SUBAPPLICATION Boot_Melden_OPC (* Station meldet ihren Start an STG1: steigende Flanke von READY ruft die Boot-Methode mit der STG-Nummer auf (ohne VT) *)
  (* Standard: 61499-2; Description: Copyright (c) 2026 Meisterschulen am Ostbahnhof This program and the accompanying materials are made available under the terms of the Eclipse Public License 2.0 which is available at https://www.eclipse.org/legal/epl-2.0/ SPDX-License-Identifier: EPL-2.0 *)
  (* Version 1.1, 2026-10-30, Franz Höpfinger, Meisterschulen am Ostbahnhof, CLIENT_1_0 (Methode) und AX_SUBSCRIBE_1 (READY) je mit Remote_Init_Retry: INITO sofort, nach INITO- (STG1 noch nicht da) neuer Versuch nach 2 s. Vorher hielt die Kette bis 60 s und der Client war danach tot (forte #1092). *)
  (* Version 1.0, 2026-10-29, Franz Höpfinger, Meisterschulen am Ostbahnhof, Neu, Gegenstueck zu Boot_Zaehler_OPC (STG1). AX_SUBSCRIBE_1 startet mit FALSE, daher gibt es nach jedem eigenen Start genau eine steigende Flanke, sobald READY von STG1 ankommt. Reconnect ohne Neustart erzeugt keine Flanke. *)
  PACKAGE MyLib::sys;
  (* Documentation:
  Start an STG1 melden
   Die Station abonniert READY von STG1. Nach dem eigenen Start steht der Wert zunächst auf FALSE; sobald TRUE von STG1 ankommt, ruft die Station einmal die Methode BOOT_MELDUNG mit ihrer Nummer NR auf. STG1 zählt die Starts (Boot_Zaehler_OPC).
  *)
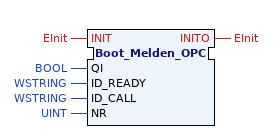
  EVENT_INPUT
    INIT : EInit; (* Initialization Request *)
  END_EVENT
  EVENT_OUTPUT
    INITO : EInit; (* Initialization Confirm *)
  END_EVENT
  VAR_INPUT
    QI : BOOL := TRUE; (* Quality Input - TRUE to enable service *)
    ID_READY : WSTRING; (* Remote-Subscribe READY von STG1 *)
    ID_CALL : WSTRING; (* Remote-Methode BOOT_MELDUNG auf STG1 *)
    NR : UINT; (* Eigene STG-Nummer (2..5) *)
  END_VAR
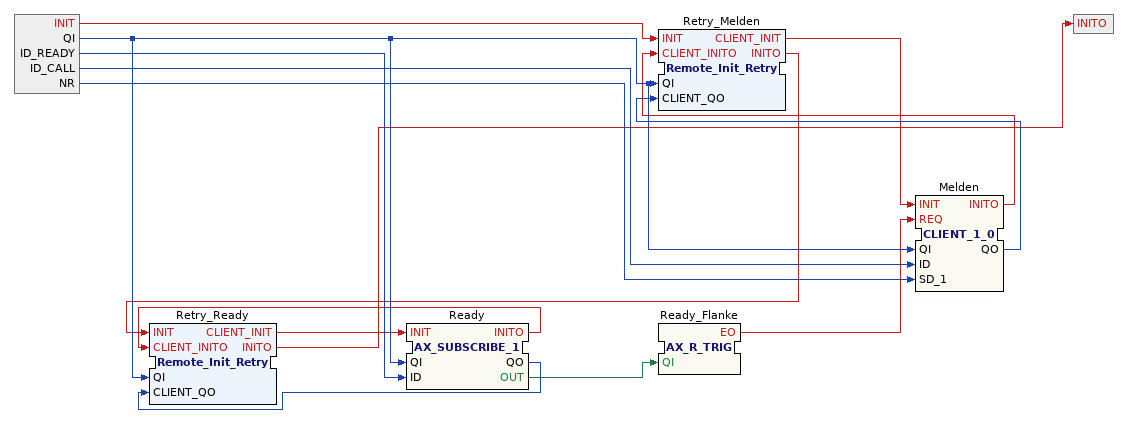
  FBS
    Melden : iec61499::net::CLIENT_1_0;
    Ready : adapter::net::AX_SUBSCRIBE_1;
    Ready_Flanke : adapter::events::unidirectional::AX_R_TRIG;
  END_FBS
  SUBAPPS
    Retry_Melden : MyLib::sys::Remote_Init_Retry;
    Retry_Ready : MyLib::sys::Remote_Init_Retry;
  END_SUBAPPS
  EVENT_CONNECTIONS
    INIT TO Retry_Melden.INIT;
    Retry_Melden.CLIENT_INIT TO Melden.INIT;
    Melden.INITO TO Retry_Melden.CLIENT_INITO;
    Retry_Melden.INITO TO Retry_Ready.INIT;
    Retry_Ready.CLIENT_INIT TO Ready.INIT;
    Ready.INITO TO Retry_Ready.CLIENT_INITO;
    Retry_Ready.INITO TO INITO;
    Ready_Flanke.EO TO Melden.REQ;
  END_CONNECTIONS
  DATA_CONNECTIONS
    QI TO Retry_Melden.QI;
    Melden.QO TO Retry_Melden.CLIENT_QO;
    QI TO Retry_Ready.QI;
    Ready.QO TO Retry_Ready.CLIENT_QO;
    QI TO Melden.QI;
    ID_CALL TO Melden.ID;
    NR TO Melden.SD_1;
    QI TO Ready.QI;
    ID_READY TO Ready.ID;
  END_CONNECTIONS
  ADAPTER_CONNECTIONS
    Ready.OUT TO Ready_Flanke.QI;
  END_CONNECTIONS
END_SUBAPPLICATION
